PROGRAM RunStudent
VAR
	LampStudent_0: LampStudent;
	ixStrobOne :BOOL;
	ixStrobTwo :BOOL;
	ixStrob: BOOL;
	LongHandshake_0: LongHandshake;
	ShortHandshake_0: ShortHandshake;
END_VAR

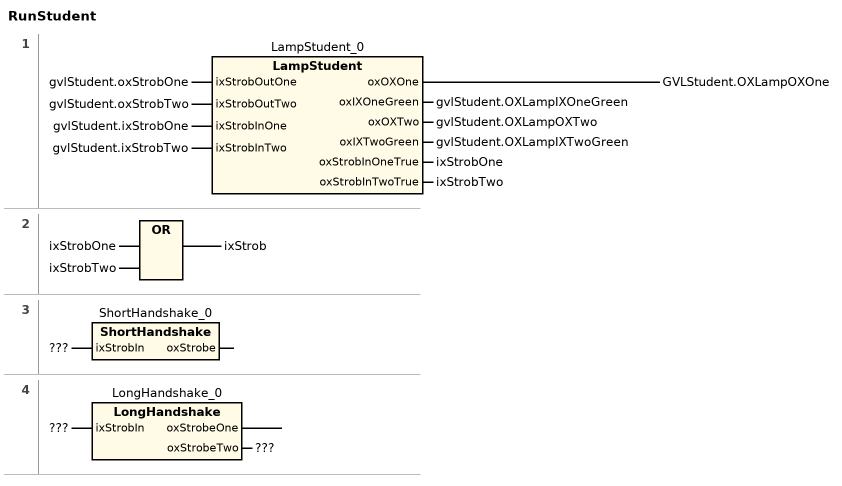
// NETWORK 1
LampStudent_0(
    ixStrobOutOne := gvlStudent.oxStrobOne,
    ixStrobOutTwo := gvlStudent.oxStrobTwo,
    ixStrobInOne := gvlStudent.ixStrobOne,
    ixStrobInTwo := gvlStudent.ixStrobTwo,
    oxIXOneGreen => gvlStudent.OXLampIXOneGreen,
    oxOXTwo => gvlStudent.OXLampOXTwo,
    oxIXTwoGreen => gvlStudent.OXLampIXTwoGreen,
    oxStrobInOneTrue => ixStrobOne,
    oxStrobInTwoTrue => ixStrobTwo); // LampStudent
GVLStudent.OXLampOXOne := LampStudent_0.oxOXOne;

// NETWORK 2
ixStrob := ixStrobOne OR ixStrobTwo;

// NETWORK 3
ShortHandshake_0(); // ShortHandshake

// NETWORK 4
LongHandshake_0(); // LongHandshake

END_PROGRAM

(* stored: Version 1.1.0.1, ProductVersion 3.1.4026.17
   POU RunStudent: Id {a6e53ef6-89cb-4074-b0db-f8344b051c13}, SpecialFunc None *)
